{region 'Documentation'}
(*!
<summary>Check that IN is less than Maximum.</summary>
<description>

All checked operands and bounds must be finite; NaN or either infinity reports Error
during active evaluation.

Numeric diagnostics use the formatter's default six significant digits; rounding affects
the message only, not the comparison.

</description>
*)
{endregion}
FUNCTION_BLOCK AssertLessThan_LReal EXTENDS AssertionBase
VAR_INPUT
    IN : LREAL; //! Actual value checked or observed by this Assertion.
    Maximum : LREAL; //! Exclusive upper bound; the actual value or count must be smaller.
END_VAR

SUPER^();

{region 'Documentation'}
(*!
<summary>Check that IN is less than Maximum.</summary>
*)
{endregion}
METHOD PROTECTED Assert
VAR
    Message : STRING(GVL_Constants.MessageLength);
    MaximumText : STRING(GVL_Constants.AssertionValueLength);
    ActualText : STRING(GVL_Constants.AssertionValueLength);
END_VAR
IF NOT EvaluationActive THEN
    RETURN;
END_IF;

IF Result = E_Result.Error THEN
    RETURN;
END_IF;

IF NOT Tc2_Utilities.LrealIsFinite(x := IN) THEN
    Error(Message := 'Assertion error: IN must be finite.');
    RETURN;
END_IF;

IF NOT Tc2_Utilities.LrealIsFinite(x := Maximum) THEN
    Error(Message := 'Assertion error: Maximum must be finite.');
    RETURN;
END_IF;

IF Result = E_Result.Failed THEN
    RETURN;
END_IF;

IF IN >= Maximum THEN
    MaximumText := CreateAssertionTextValue_LReal(Value := Maximum);
    ActualText := CreateAssertionTextValue_LReal(Value := IN);
    Message := CONCAT('Assertion failed: value is not less than maximum. Maximum = ',
        MaximumText);
    Message := CONCAT(Message, ', Actual = ');
    Message := CONCAT(Message, ActualText);
    Message := CONCAT(Message, '.');
    Fail(Message := Message);
    RETURN;
END_IF;

Pass();
END_METHOD

END_FUNCTION_BLOCK

(* stored: Version 1.1.0.1
   POU AssertLessThan_LReal: Id {09d35e1b-c1e7-4883-aba9-c9414d7ce58f}, SpecialFunc None
   Folder Internal: Id {b56cf2e4-aeab-4ec0-89be-097e7785762d}
   Method Assert: Id {4e071cc3-2b7c-497e-b663-b8aa559b0ecc} *)
